{attribute 'qualified_only'}
{attribute 'strict'}
TYPE E_Tank_Name :
(
	enum_member := 0,
	
	//CIP
	T91,
	T92,
	T93,
	T94,
	
	//Marinade
	T1,
	T2,
	
	//Color
	T3,
	T4,
	
	last
	
);
END_TYPE

(* stored: Version 1.1.0.1, ProductVersion 3.1.4024.12
   EnumerationTextList E_Tank_Name: Id {a6265d94-a280-4b35-91b4-69cbc2a882b9} *)
